Fanuc KAREL source: KT00540.KL

PROGRAM KT00540
%NOLOCKGROUP
VAR
  P1: JOINTPOS
  P2: XYZWPR
  OUT: XYZWPR
BEGIN
    P2.Y = 2.0
  OUT = P1 : P2
END KT00540
